(* IEC 61131-3 sources: llm-plc-st-eval/codesys/dobles/I2, 6 files *)

(* ---- 01_Correcta.st ---- *)
(* DOBLE DE PRUEBA I2/Correcta - NO ES CORPUS. Esperado: veredicto 1 *)
FUNCTION_BLOCK FB_Llenado
VAR_INPUT
    nivelAlto : BOOL;
    nivelBajo : BOOL;
    btnInicio : BOOL;
    btnParo : BOOL;
END_VAR
VAR_OUTPUT
    vLlenado : BOOL;
    motorMezcla : BOOL;
    vDescarga : BOOL;
END_VAR
VAR
    tAhora : TIME;
    tPrev : TIME;
    dScan : TIME;
    init : BOOL;
    estado : INT;
    t : TIME;
END_VAR
tAhora := TIME();
IF NOT init THEN
    tPrev := tAhora;
    init := TRUE;
END_IF
dScan := tAhora - tPrev;
tPrev := tAhora;
IF btnParo THEN
    vLlenado := FALSE; motorMezcla := FALSE; vDescarga := FALSE;
    estado := 0;
    t := T#0S;
ELSE
    CASE estado OF
        0:
            vLlenado := FALSE; motorMezcla := FALSE; vDescarga := FALSE;
            IF btnInicio THEN estado := 1; END_IF
        1:
            vLlenado := TRUE; motorMezcla := FALSE; vDescarga := FALSE;
            IF nivelAlto THEN estado := 2; t := T#0S; END_IF
        2:
            vLlenado := FALSE; motorMezcla := TRUE; vDescarga := FALSE;
            t := t + dScan;
            IF t >= T#60S THEN estado := 3; END_IF
    ELSE
            vLlenado := FALSE; motorMezcla := FALSE; vDescarga := TRUE;
            IF nivelBajo THEN estado := 0; END_IF
    END_CASE
END_IF
END_FUNCTION_BLOCK

(* ---- 02_MezclaCorta.st ---- *)
(* DOBLE DE PRUEBA I2/MezclaCorta - NO ES CORPUS. Esperado: veredicto 2, falla en el paso 3 *)
FUNCTION_BLOCK FB_Llenado
VAR_INPUT
    nivelAlto : BOOL;
    nivelBajo : BOOL;
    btnInicio : BOOL;
    btnParo : BOOL;
END_VAR
VAR_OUTPUT
    vLlenado : BOOL;
    motorMezcla : BOOL;
    vDescarga : BOOL;
END_VAR
VAR
    tAhora : TIME;
    tPrev : TIME;
    dScan : TIME;
    init : BOOL;
    estado : INT;
    t : TIME;
END_VAR
tAhora := TIME();
IF NOT init THEN
    tPrev := tAhora;
    init := TRUE;
END_IF
dScan := tAhora - tPrev;
tPrev := tAhora;
IF btnParo THEN
    vLlenado := FALSE; motorMezcla := FALSE; vDescarga := FALSE;
    estado := 0;
    t := T#0S;
ELSE
    CASE estado OF
        0:
            vLlenado := FALSE; motorMezcla := FALSE; vDescarga := FALSE;
            IF btnInicio THEN estado := 1; END_IF
        1:
            vLlenado := TRUE; motorMezcla := FALSE; vDescarga := FALSE;
            IF nivelAlto THEN estado := 2; t := T#0S; END_IF
        2:
            vLlenado := FALSE; motorMezcla := TRUE; vDescarga := FALSE;
            t := t + dScan;
            IF t >= T#30S THEN estado := 3; END_IF
    ELSE
            vLlenado := FALSE; motorMezcla := FALSE; vDescarga := TRUE;
            IF nivelBajo THEN estado := 0; END_IF
    END_CASE
END_IF
END_FUNCTION_BLOCK

(* ---- 03_SaltaMezcla.st ---- *)
(* DOBLE DE PRUEBA I2/SaltaMezcla - NO ES CORPUS. Esperado: veredicto 2, falla en el paso 2 *)
FUNCTION_BLOCK FB_Llenado
VAR_INPUT
    nivelAlto : BOOL;
    nivelBajo : BOOL;
    btnInicio : BOOL;
    btnParo : BOOL;
END_VAR
VAR_OUTPUT
    vLlenado : BOOL;
    motorMezcla : BOOL;
    vDescarga : BOOL;
END_VAR
VAR
    tAhora : TIME;
    tPrev : TIME;
    dScan : TIME;
    init : BOOL;
    estado : INT;
    t : TIME;
END_VAR
tAhora := TIME();
IF NOT init THEN
    tPrev := tAhora;
    init := TRUE;
END_IF
dScan := tAhora - tPrev;
tPrev := tAhora;
IF btnParo THEN
    vLlenado := FALSE; motorMezcla := FALSE; vDescarga := FALSE;
    estado := 0;
    t := T#0S;
ELSE
    CASE estado OF
        0:
            vLlenado := FALSE; motorMezcla := FALSE; vDescarga := FALSE;
            IF btnInicio THEN estado := 1; END_IF
        1:
            vLlenado := TRUE; motorMezcla := FALSE; vDescarga := FALSE;
            IF nivelAlto THEN estado := 3; t := T#0S; END_IF
        2:
            vLlenado := FALSE; motorMezcla := TRUE; vDescarga := FALSE;
            t := t + dScan;
            IF t >= T#60S THEN estado := 3; END_IF
    ELSE
            vLlenado := FALSE; motorMezcla := FALSE; vDescarga := TRUE;
            IF nivelBajo THEN estado := 0; END_IF
    END_CASE
END_IF
END_FUNCTION_BLOCK

(* ---- 04_ParoNoSeguro.st ---- *)
(* DOBLE DE PRUEBA I2/ParoNoSeguro - NO ES CORPUS. Esperado: veredicto 2, falla en el paso 7 *)
FUNCTION_BLOCK FB_Llenado
VAR_INPUT
    nivelAlto : BOOL;
    nivelBajo : BOOL;
    btnInicio : BOOL;
    btnParo : BOOL;
END_VAR
VAR_OUTPUT
    vLlenado : BOOL;
    motorMezcla : BOOL;
    vDescarga : BOOL;
END_VAR
VAR
    tAhora : TIME;
    tPrev : TIME;
    dScan : TIME;
    init : BOOL;
    estado : INT;
    t : TIME;
END_VAR
tAhora := TIME();
IF NOT init THEN
    tPrev := tAhora;
    init := TRUE;
END_IF
dScan := tAhora - tPrev;
tPrev := tAhora;
IF btnParo THEN
    estado := 0;
    t := T#0S;
ELSE
    CASE estado OF
        0:
            vLlenado := FALSE; motorMezcla := FALSE; vDescarga := FALSE;
            IF btnInicio THEN estado := 1; END_IF
        1:
            vLlenado := TRUE; motorMezcla := FALSE; vDescarga := FALSE;
            IF nivelAlto THEN estado := 2; t := T#0S; END_IF
        2:
            vLlenado := FALSE; motorMezcla := TRUE; vDescarga := FALSE;
            t := t + dScan;
            IF t >= T#60S THEN estado := 3; END_IF
    ELSE
            vLlenado := FALSE; motorMezcla := FALSE; vDescarga := TRUE;
            IF nivelBajo THEN estado := 0; END_IF
    END_CASE
END_IF
END_FUNCTION_BLOCK

(* ---- 05_ParoSoloEnLlenado.st ---- *)
(* DOBLE DE PRUEBA I2/ParoSoloEnLlenado - NO ES CORPUS. Esperado: veredicto 2, falla en el paso 10 *)
FUNCTION_BLOCK FB_Llenado
VAR_INPUT
    nivelAlto : BOOL;
    nivelBajo : BOOL;
    btnInicio : BOOL;
    btnParo : BOOL;
END_VAR
VAR_OUTPUT
    vLlenado : BOOL;
    motorMezcla : BOOL;
    vDescarga : BOOL;
END_VAR
VAR
    tAhora : TIME;
    tPrev : TIME;
    dScan : TIME;
    init : BOOL;
    estado : INT;
    t : TIME;
END_VAR
tAhora := TIME();
IF NOT init THEN
    tPrev := tAhora;
    init := TRUE;
END_IF
dScan := tAhora - tPrev;
tPrev := tAhora;
IF btnParo AND estado <> 2 THEN
    vLlenado := FALSE; motorMezcla := FALSE; vDescarga := FALSE;
    estado := 0;
    t := T#0S;
ELSE
    CASE estado OF
        0:
            vLlenado := FALSE; motorMezcla := FALSE; vDescarga := FALSE;
            IF btnInicio THEN estado := 1; END_IF
        1:
            vLlenado := TRUE; motorMezcla := FALSE; vDescarga := FALSE;
            IF nivelAlto THEN estado := 2; t := T#0S; END_IF
        2:
            vLlenado := FALSE; motorMezcla := TRUE; vDescarga := FALSE;
            t := t + dScan;
            IF t >= T#60S THEN estado := 3; END_IF
    ELSE
            vLlenado := FALSE; motorMezcla := FALSE; vDescarga := TRUE;
            IF nivelBajo THEN estado := 0; END_IF
    END_CASE
END_IF
END_FUNCTION_BLOCK

(* ---- 06_NoRearranca.st ---- *)
(* DOBLE DE PRUEBA I2/NoRearranca - NO ES CORPUS. Esperado: veredicto 2, falla en el paso 8 *)
FUNCTION_BLOCK FB_Llenado
VAR_INPUT
    nivelAlto : BOOL;
    nivelBajo : BOOL;
    btnInicio : BOOL;
    btnParo : BOOL;
END_VAR
VAR_OUTPUT
    vLlenado : BOOL;
    motorMezcla : BOOL;
    vDescarga : BOOL;
END_VAR
VAR
    tAhora : TIME;
    tPrev : TIME;
    dScan : TIME;
    init : BOOL;
    estado : INT;
    t : TIME;
    bloqueado : BOOL;
END_VAR
tAhora := TIME();
IF NOT init THEN
    tPrev := tAhora;
    init := TRUE;
END_IF
dScan := tAhora - tPrev;
tPrev := tAhora;
IF btnParo THEN
    vLlenado := FALSE; motorMezcla := FALSE; vDescarga := FALSE;
    estado := 0;
    t := T#0S;
    bloqueado := TRUE;
ELSE
    IF bloqueado THEN
        vLlenado := FALSE; motorMezcla := FALSE; vDescarga := FALSE;
    ELSE
        CASE estado OF
            0:
                vLlenado := FALSE; motorMezcla := FALSE; vDescarga := FALSE;
                IF btnInicio THEN estado := 1; END_IF
            1:
                vLlenado := TRUE; motorMezcla := FALSE; vDescarga := FALSE;
                IF nivelAlto THEN estado := 2; t := T#0S; END_IF
            2:
                vLlenado := FALSE; motorMezcla := TRUE; vDescarga := FALSE;
                t := t + dScan;
                IF t >= T#60S THEN estado := 3; END_IF
        ELSE
                vLlenado := FALSE; motorMezcla := FALSE; vDescarga := TRUE;
                IF nivelBajo THEN estado := 0; END_IF
        END_CASE
    END_IF
END_IF
END_FUNCTION_BLOCK
